(* IEC 61131-3 sources: plc-process-lib/tests/POUs/Suites/FB_Common_Test, 10 files *)

(* ---- CfgDefaultsMatchContract.method.decl.st ---- *)
// Значения Cfg по умолчанию — по контракту (на них опирается генератор: экземпляр без строки
// конфигурации корректен). Инициализатор элемента массива (ePriority := ...) оставляет прочим
// полям умолчания ST_AlarmCfg (проверка R9 контракта для DUT).
METHOD PRIVATE CfgDefaultsMatchContract
VAR
    stAlm : ST_AlarmCfg;           // умолчания ST_AlarmCfg
    stSlot : ST_AlarmCfg;          // копия элемента astAlarm[i]
    stLim : ST_AiLimitCfg;         // копия элемента astLimit[i]
    stAi  : ST_AnalogInputCfg;
    stDi  : ST_DigitalInputCfg;
    stMot : ST_MotorCfg;
    stVlv : ST_ValveCfg;
    stCv  : ST_ControlValveCfg;
    stPid : ST_PidCfg;
END_VAR

(* ---- InterfaceRefsDefaultToNull.method.decl.st ---- *)
// Интерфейсные ссылки до присваивания — 0 (так их проверяют ФБ: itfTime <> 0); цепочка EXTENDS
// I_MotorVfd → I_Motor → I_Device → I_AlarmSource допускает приведение вверх.
METHOD PRIVATE InterfaceRefsDefaultToNull
VAR
    itfTime     : I_TimeSource;
    itfAlarm    : I_Alarm;
    itfSource   : I_AlarmSource;
    itfDevice   : I_Device;
    itfMotor    : I_Motor;
    itfMotorVfd : I_MotorVfd;
    itfSink     : I_AlarmSink;
END_VAR

(* ---- SizeOfAlarmCfgIs16.method.decl.st ---- *)
// SIZEOF(ST_AlarmCfg) = 16 (зонд Q14 контракта) и SIZEOF(ST_AiLimitCfg) = 20: элементы массивов
// astAlarm и astLimit в persistent-данных. Источник: tools/reference/common.py, сценарий cfg_sizes.
METHOD PRIVATE SizeOfAlarmCfgIs16
VAR
    stAlm : ST_AlarmCfg;           // параметры тревоги
    stLim : ST_AiLimitCfg;         // параметры уставки
END_VAR

(* ---- SizeOfCfgMatchesReference.method.decl.st ---- *)
// SIZEOF структур Cfg — по расчёту раскладки (Control Win V3 32 бит). Cfg лежат в Persistent
// Variables приложения: изменение типа переинициализирует уставки (A-13), тест ловит его.
// Источник: tools/reference/common.py, сценарий cfg_sizes.
METHOD PRIVATE SizeOfCfgMatchesReference
VAR
    stAi  : ST_AnalogInputCfg;
    stDi  : ST_DigitalInputCfg;
    stMot : ST_MotorCfg;
    stVfd : ST_VfdCfg;
    stVlv : ST_ValveCfg;
    stCv  : ST_ControlValveCfg;
    stPid : ST_PidCfg;
END_VAR

(* ---- SizeOfCmdMatchesReference.method.decl.st ---- *)
// SIZEOF структур команд HMI/SCADA (GVL_Hmi приложения). Источник: tools/reference/common.py, сценарий cmd_sizes.
METHOD PRIVATE SizeOfCmdMatchesReference
VAR
    stDev : ST_DeviceCmd;          // общий заголовок
    stAi  : ST_AnalogInputCmd;
    stDi  : ST_DigitalInputCmd;
    stMot : ST_MotorCmd;
    stVlv : ST_ValveCmd;
    stCv  : ST_ControlValveCmd;
    stPid : ST_PidCmd;
END_VAR

(* ---- SizeOfDeviceRetainIs36.method.decl.st ---- *)
// SIZEOF(ST_DeviceRetain) = 36 на Control Win V3 32 бит (зонд P17 контракта).
METHOD PRIVATE SizeOfDeviceRetainIs36
VAR
    stRetain : ST_DeviceRetain;    // энергонезависимые данные устройства
END_VAR

(* ---- SizeOfStsMatchesRegisterMap.method.decl.st ---- *)
// SIZEOF семи структур состояния — таблица 4.6 контракта (карта регистров Modbus = порядок полей,
// скрытого выравнивания нет). Источник: таблица 4.6 и tools/reference/common.py, сценарий sts_sizes.
METHOD PRIVATE SizeOfStsMatchesRegisterMap
VAR
    stDev : ST_DeviceSts;          // общий заголовок
    stAi  : ST_AnalogInputSts;
    stDi  : ST_DigitalInputSts;
    stMot : ST_MotorSts;           // и для FB_MotorVfd
    stVlv : ST_ValveSts;
    stCv  : ST_ControlValveSts;
    stPid : ST_PidSts;
END_VAR

(* ---- StsRetainDefaultsMatchContract.method.decl.st ---- *)
// Умолчания общего заголовка и энергонезависимых данных: до первого вызова eMode = Manual,
// eNe107 = CheckFunction («не проверено»), тип None; дистанционный режим в Retain — Manual.
// Вложенный заголовок stCommon сохраняет свои умолчания.
METHOD PRIVATE StsRetainDefaultsMatchContract
VAR
    stDev    : ST_DeviceSts;       // общий заголовок
    stMot    : ST_MotorSts;        // вложенный заголовок
    stRetain : ST_DeviceRetain;    // энергонезависимые данные
END_VAR

(* ---- TestSinkRecordsEventsInOrder.method.decl.st ---- *)
// FB_TestSink через PL.GVL_Lib.itfAlarmSink (как его вызывает FB_Alarm): события по порядку,
// Last и GetEvent, кольцо на 32 события (33 события — остаются 32 последних), Clear. Приёмник
// возвращается в 0 до конца теста.
METHOD PRIVATE TestSinkRecordsEventsInOrder
VAR
    fbSink    : FB_TestSink;       // приёмник под тестом
    stEv1     : ST_AlarmEvent;     // первое событие
    stEv2     : ST_AlarmEvent;     // второе событие
    stGot     : ST_AlarmEvent;     // прочитанное событие
    xAccepted : BOOL;              // ответ приёмника
    uiEvent   : UINT;              // номер события в цикле
END_VAR

(* ---- TestSinkRecordsEventsInOrder.method.impl.st ---- *)
coUnit.TEST('Common_TestSink_RecordsEventsInOrder');

stEv1.udiId := 121;
stEv1.ePriority := E_AlarmPriority.High;
stEv1.eOldState := E_AlarmState.Normal;
stEv1.eNewState := E_AlarmState.ActiveUnack;
stEv1.eReason := E_AlarmEventReason.Activated;
stEv1.ltTime := LTIME#1H;
stEv1.rValue := 4.5;
stEv2 := stEv1;
stEv2.udiId := 122;
stEv2.eOldState := E_AlarmState.ActiveUnack;
stEv2.eNewState := E_AlarmState.ActiveAck;
stEv2.eReason := E_AlarmEventReason.Acked;
stEv2.ltTime := LTIME#2H;

GVL_Lib.itfAlarmSink := fbSink;
xAccepted := GVL_Lib.itfAlarmSink.OnAlarmEvent(stEvent := stEv1);
GVL_Lib.itfAlarmSink.OnAlarmEvent(stEvent := stEv2);
GVL_Lib.itfAlarmSink := 0;                                     // приёмник — снова 0

AssertTrue(Condition := xAccepted, Message := 'sink accepts the event');
AssertEquals_UINT(Expected := 2, Actual := fbSink.Count, Message := 'two events recorded');
stGot := fbSink.Last;
AssertEquals_UDINT(Expected := 122, Actual := stGot.udiId, Message := 'last event is the second one');
AssertTrue(Condition := stGot.eReason = E_AlarmEventReason.Acked, Message := 'last event reason Acked');
stGot := fbSink.GetEvent(uiBack := 1);
AssertEquals_UDINT(Expected := 121, Actual := stGot.udiId, Message := 'previous event is the first one');
AssertEquals_LTIME(Expected := LTIME#1H, Actual := stGot.ltTime, Message := 'event time stamp kept');
AssertEquals_REAL(Expected := 4.5, Actual := stGot.rValue, Delta := 0.0, Message := 'event value kept');
AssertTrue(Condition := GVL_Lib.itfAlarmSink = 0, Message := 'library sink restored to 0');

FOR uiEvent := 1 TO 33 DO
    stEv1.udiId := 1000 + uiEvent;
    fbSink.OnAlarmEvent(stEvent := stEv1);
END_FOR
AssertEquals_UINT(Expected := 35, Actual := fbSink.Count, Message := 'all events counted');
stGot := fbSink.Last;
AssertEquals_UDINT(Expected := 1033, Actual := stGot.udiId, Message := 'last of 33 events');
stGot := fbSink.GetEvent(uiBack := 31);
AssertEquals_UDINT(Expected := 1002, Actual := stGot.udiId, Message := 'the ring keeps the last 32 events');
stGot := fbSink.GetEvent(uiBack := 32);
AssertEquals_UDINT(Expected := 0, Actual := stGot.udiId, Message := 'older events are gone: empty event');

fbSink.Clear();
AssertEquals_UINT(Expected := 0, Actual := fbSink.Count, Message := 'Clear forgets all events');
stGot := fbSink.Last;
AssertEquals_UDINT(Expected := 0, Actual := stGot.udiId, Message := 'no last event after Clear');

coUnit.TEST_FINISHED();
